(* Tests trace and span identifier generation.

   A generator fills its ring from the operating system guid service over ADS, so a fresh one
   has nothing to hand out until tick has been pumped for a few cycles. Every test that needs
   identifiers waits for that first refill before asserting anything about the bytes it gets
   back.

   Each test declares its generator in its own VAR_INST, next to the state machine that pumps
   it, so the ring a test reasons about is written down where the test reads it rather than in
   a list on the suite. Ring sizes are therefore chosen per test: most take a ring far larger
   than they draw from, so the seam never comes into it, while the wrap and capacity tests
   deliberately take the smallest ring the configuration allows, because a ring that small is
   the only one a test can drain often enough to lap. *)
FUNCTION_BLOCK FB_TestIdGenerator EXTENDS FB_TestSuite

THIS^.testRejectsInvalidConfiguration();
THIS^.testFailsBeforeTheFirstRefill();
THIS^.testGeneratesUniqueTraceIds();
THIS^.testGeneratesUniqueSpanIds();
THIS^.testDrawsAcrossTheWrap();
THIS^.testHonorsConfiguredCapacity();
THIS^.testGeneratesThroughTheBaseReference();
THIS^.testSeparateGeneratorsDoNotCollide();

(* TRUE when every byte in the buffer is zero, which is the identifier OTLP reads as absent. *)
METHOD _isZero : BOOL
VAR_INPUT
	pBytes: POINTER TO BYTE;
	nBytes: UDINT;
END_VAR
VAR
	_idx: UDINT;
END_VAR
_isZero := TRUE;

IF (pBytes = 0) OR_ELSE (nBytes = 0) THEN
	RETURN;
END_IF

FOR _idx := 0 TO nBytes - 1 DO
	IF pBytes[_idx] <> 0 THEN
		_isZero := FALSE;
		RETURN;
	END_IF
END_FOR
END_METHOD

(* Exercises the seam. A thirty two byte ring cannot hold eight identifiers at once, so the
   draws are spread over cycles and the read point laps the ring several times.

   Taking sixteen bytes and then eight moves the read point by twenty four, which lands it on
   every eight byte alignment in turn: some trace draws stop short of the end of the ring, one
   ends exactly on it, and one starts near the end and has to be stitched from both sides. A
   stitch that copied the wrong end, or re-read bytes already handed out, shows up here as a
   repeat among the samples. *)
METHOD testDrawsAcrossTheWrap : REFERENCE TO FB_Test

VAR CONSTANT
	MAX_CYCLES: UDINT := 60000;
	SAMPLES: UDINT := 8;
END_VAR

VAR_INST
	_generator: FB_IdGenerator(nTraceIds := 1, nSpanIds := 1);  // 24 bytes, which FB_Init rounds up to 32
	_cycles: UDINT;
	_state: USINT;
	_traceIdx: UDINT;
	_spanIdx: UDINT;
	_traceSamples: ARRAY [0..7, 0..15] OF BYTE;  // held across cycles, unlike the other suites
	_spanSamples: ARRAY [0..7, 0..7] OF BYTE;
END_VAR

VAR
	traceId: FB_TraceId;
	spanId: FB_SpanId;
	failureReason: E_IdGenFailureReason;
	tickSucceeded: BOOL;
	_i: UDINT;
	_j: UDINT;
END_VAR
TcUnit.TEST('testDrawsAcrossTheWrap');
	CASE _state OF
		0: // take whatever the ring can serve this cycle, however many laps that takes
			tickSucceeded := _generator.tick(failureReason=>failureReason);
			_cycles := _cycles + 1;
			IF NOT tickSucceeded THEN
				THIS^.AssertTrue(FALSE, 'Expected the guid service to refill the ring without error');
				_state := 255;
				TcUnit.TEST_FINISHED();
				RETURN;
			END_IF

			IF (_traceIdx < SAMPLES) AND_THEN _generator.generateTraceId(traceId:=traceId, failureReason=>failureReason) THEN
				MEMCPY(ADR(_traceSamples[_traceIdx, 0]), ADR(traceId.bytes), SIZEOF(traceId.bytes));
				_traceIdx := _traceIdx + 1;
			END_IF

			IF (_spanIdx < SAMPLES) AND_THEN _generator.generateSpanId(spanId:=spanId, failureReason=>failureReason) THEN
				MEMCPY(ADR(_spanSamples[_spanIdx, 0]), ADR(spanId.bytes), SIZEOF(spanId.bytes));
				_spanIdx := _spanIdx + 1;
			END_IF

			IF (_traceIdx >= SAMPLES) AND (_spanIdx >= SAMPLES) THEN
				_state := 10;
			ELSIF _cycles > MAX_CYCLES THEN
				THIS^.AssertTrue(FALSE, 'Expected a ring small enough to wrap to hand out its identifiers within MAX_CYCLES');
				_state := 255;
				TcUnit.TEST_FINISHED();
			END_IF
			RETURN;

		10:
			FOR _i := 0 TO 7 DO
				THIS^.AssertFalse(
					THIS^._isZero(pBytes:=ADR(_traceSamples[_i, 0]), nBytes:=TO_UDINT(SIZEOF(traceId.bytes))),
					'Expected no trace id drawn from a wrapping ring to be all zeroes'
				);
				THIS^.AssertFalse(
					THIS^._isZero(pBytes:=ADR(_spanSamples[_i, 0]), nBytes:=TO_UDINT(SIZEOF(spanId.bytes))),
					'Expected no span id drawn from a wrapping ring to be all zeroes'
				);

				FOR _j := 0 TO 7 DO
					IF _i <> _j THEN
						THIS^.AssertTrue(
							MEMCMP(ADR(_traceSamples[_i, 0]), ADR(_traceSamples[_j, 0]), SIZEOF(traceId.bytes)) <> 0,
							'Expected every trace id to differ, including the one stitched across the wrap'
						);
						THIS^.AssertTrue(
							MEMCMP(ADR(_spanSamples[_i, 0]), ADR(_spanSamples[_j, 0]), SIZEOF(spanId.bytes)) <> 0,
							'Expected every span id to differ, including the ones taken either side of the wrap'
						);
					END_IF
				END_FOR
			END_FOR

			_state := 255;
			TcUnit.TEST_FINISHED();
			RETURN;
	END_CASE
END_METHOD

(* A generator that has never been ticked holds no bytes. It has to say so, because the only
   thing it could hand out instead is the all zero identifier OTLP reads as absent. *)
METHOD testFailsBeforeTheFirstRefill : REFERENCE TO FB_Test

VAR_INST
	_generator: FB_IdGenerator(nTraceIds := 16, nSpanIds := 16);  // deliberately never ticked, so it stays empty
	_state: USINT;
END_VAR

VAR
	traceId: FB_TraceId;
	spanId: FB_SpanId;
	failureReason: E_IdGenFailureReason;
	success: BOOL;
END_VAR
TcUnit.TEST('testFailsBeforeTheFirstRefill');
	CASE _state OF
		0:
			THIS^.AssertTrue(_generator.configValid, 'Expected a generator with a ring to report a valid configuration');

			success := _generator.generateTraceId(traceId:=traceId, failureReason=>failureReason);
			THIS^.AssertFalse(success, 'Expected trace id generation to fail before the first refill');
			THIS^.AssertEquals_UDINT(
				TO_UDINT(E_IdGenFailureReason.NO_IDENTIFIERS_AVAILABLE),
				TO_UDINT(failureReason),
				'Expected an empty ring to report NO_IDENTIFIERS_AVAILABLE'
			);
			THIS^.AssertTrue(
				THIS^._isZero(pBytes:=ADR(traceId.bytes), nBytes:=TO_UDINT(SIZEOF(traceId.bytes))),
				'Expected a failed draw to leave the trace id untouched'
			);

			success := _generator.generateSpanId(spanId:=spanId, failureReason=>failureReason);
			THIS^.AssertFalse(success, 'Expected span id generation to fail before the first refill');
			THIS^.AssertEquals_UDINT(
				TO_UDINT(E_IdGenFailureReason.NO_IDENTIFIERS_AVAILABLE),
				TO_UDINT(failureReason),
				'Expected an empty ring to report NO_IDENTIFIERS_AVAILABLE'
			);
			THIS^.AssertTrue(
				THIS^._isZero(pBytes:=ADR(spanId.bytes), nBytes:=TO_UDINT(SIZEOF(spanId.bytes))),
				'Expected a failed draw to leave the span id untouched'
			);

			_state := 255;
			TcUnit.TEST_FINISHED();
	END_CASE
END_METHOD

(* Callers hold the generator as REFERENCE TO FB_IdGenerator_Base, so the abstract methods have
   to dispatch to the concrete ring. *)
METHOD testGeneratesThroughTheBaseReference : REFERENCE TO FB_Test

VAR CONSTANT
	MAX_CYCLES: UDINT := 60000;
END_VAR

VAR_INST
	_generator: FB_IdGenerator(nTraceIds := 16, nSpanIds := 16);
	_cycles: UDINT;
	_state: USINT;
END_VAR

VAR
	base: REFERENCE TO FB_IdGenerator_Base;
	traceId: FB_TraceId;
	spanId: FB_SpanId;
	failureReason: E_IdGenFailureReason;
	tickSucceeded: BOOL;
	success: BOOL;
END_VAR
TcUnit.TEST('testGeneratesThroughTheBaseReference');
	base REF= _generator;
	CASE _state OF
		0:
			THIS^.AssertTrue(__ISVALIDREF(base), 'Expected the base reference to be valid');
			_state := 10;
			RETURN;

		10: // pump through the base reference until the first refill lands
			tickSucceeded := base.tick(failureReason=>failureReason);
			_cycles := _cycles + 1;
			IF NOT tickSucceeded THEN
				THIS^.AssertTrue(FALSE, 'Expected tick to dispatch to the concrete generator without error');
				_state := 255;
				TcUnit.TEST_FINISHED();
				RETURN;
			END_IF

			success := base.generateTraceId(traceId:=traceId, failureReason=>failureReason);
			IF NOT success THEN
				IF _cycles > MAX_CYCLES THEN
					THIS^.AssertTrue(FALSE, 'Expected identifiers through the base reference within MAX_CYCLES');
					_state := 255;
					TcUnit.TEST_FINISHED();
				END_IF
				RETURN;
			END_IF

			THIS^.AssertFalse(
				THIS^._isZero(pBytes:=ADR(traceId.bytes), nBytes:=TO_UDINT(SIZEOF(traceId.bytes))),
				'Expected a non zero trace id through the base reference'
			);

			success := base.generateSpanId(spanId:=spanId, failureReason=>failureReason);
			THIS^.AssertTrue(success, 'Expected generateSpanId to dispatch to the concrete generator');
			THIS^.AssertFalse(
				THIS^._isZero(pBytes:=ADR(spanId.bytes), nBytes:=TO_UDINT(SIZEOF(spanId.bytes))),
				'Expected a non zero span id through the base reference'
			);

			_state := 255;
			TcUnit.TEST_FINISHED();
			RETURN;
	END_CASE
END_METHOD

(* The same requirement as for trace ids. A span id handed out twice makes two spans in the
   same trace indistinguishable. *)
METHOD testGeneratesUniqueSpanIds : REFERENCE TO FB_Test

VAR CONSTANT
	MAX_CYCLES: UDINT := 60000;
END_VAR

VAR_INST
	_generator: FB_IdGenerator(nTraceIds := 16, nSpanIds := 16);  // 384 bytes, so eight samples come out of one fill
	_cycles: UDINT;
	_state: USINT;
END_VAR

VAR
	spanId: FB_SpanId;
	samples: ARRAY [0..7, 0..7] OF BYTE;
	failureReason: E_IdGenFailureReason;
	tickSucceeded: BOOL;
	success: BOOL;
	_i: UDINT;
	_j: UDINT;
END_VAR
TcUnit.TEST('testGeneratesUniqueSpanIds');
	CASE _state OF
		0: // wait for the first refill before drawing the samples
			tickSucceeded := _generator.tick(failureReason=>failureReason);
			_cycles := _cycles + 1;
			IF NOT tickSucceeded THEN
				THIS^.AssertTrue(FALSE, 'Expected the guid service to refill the ring without error');
				_state := 255;
				TcUnit.TEST_FINISHED();
				RETURN;
			END_IF

			IF _generator.generateSpanId(spanId:=spanId, failureReason=>failureReason) THEN
				_state := 10;
			ELSIF _cycles > MAX_CYCLES THEN
				THIS^.AssertTrue(FALSE, 'Expected the first ring of span ids within MAX_CYCLES');
				_state := 255;
				TcUnit.TEST_FINISHED();
			END_IF
			RETURN;

		10: // a full ring holds forty eight span ids, so all eight samples come out of one fill
			FOR _i := 0 TO 7 DO
				success := _generator.generateSpanId(spanId:=spanId, failureReason=>failureReason);
				THIS^.AssertTrue(success, 'Expected every span id draw from a filled ring to succeed');
				THIS^.AssertEquals_UDINT(
					TO_UDINT(E_IdGenFailureReason.NA),
					TO_UDINT(failureReason),
					'Expected no failure reason alongside a successful draw'
				);
				THIS^.AssertFalse(
					THIS^._isZero(pBytes:=ADR(spanId.bytes), nBytes:=TO_UDINT(SIZEOF(spanId.bytes))),
					'Expected no span id to be all zeroes'
				);
				MEMCPY(ADR(samples[_i, 0]), ADR(spanId.bytes), SIZEOF(spanId.bytes));
			END_FOR

			FOR _i := 0 TO 7 DO
				FOR _j := 0 TO 7 DO
					IF _i <> _j THEN
						THIS^.AssertTrue(
							MEMCMP(ADR(samples[_i, 0]), ADR(samples[_j, 0]), SIZEOF(spanId.bytes)) <> 0,
							'Expected every span id to differ from every other'
						);
					END_IF
				END_FOR
			END_FOR

			_state := 255;
			TcUnit.TEST_FINISHED();
			RETURN;
	END_CASE
END_METHOD

(* Every draw has to be its own bytes. A trace id handed out twice merges two unrelated traces
   at the collector, which is worse than no trace at all. *)
METHOD testGeneratesUniqueTraceIds : REFERENCE TO FB_Test

VAR CONSTANT
	MAX_CYCLES: UDINT := 60000;
END_VAR

VAR_INST
	_generator: FB_IdGenerator(nTraceIds := 16, nSpanIds := 16);  // 384 bytes, so eight samples come out of one fill
	_cycles: UDINT;
	_state: USINT;
END_VAR

VAR
	traceId: FB_TraceId;
	samples: ARRAY [0..7, 0..15] OF BYTE;
	failureReason: E_IdGenFailureReason;
	tickSucceeded: BOOL;
	success: BOOL;
	_i: UDINT;
	_j: UDINT;
END_VAR
TcUnit.TEST('testGeneratesUniqueTraceIds');
	CASE _state OF
		0: // wait for the first refill before drawing the samples
			tickSucceeded := _generator.tick(failureReason=>failureReason);
			_cycles := _cycles + 1;
			IF NOT tickSucceeded THEN
				THIS^.AssertTrue(FALSE, 'Expected the guid service to refill the ring without error');
				_state := 255;
				TcUnit.TEST_FINISHED();
				RETURN;
			END_IF

			IF _generator.generateTraceId(traceId:=traceId, failureReason=>failureReason) THEN
				_state := 10;
			ELSIF _cycles > MAX_CYCLES THEN
				THIS^.AssertTrue(FALSE, 'Expected the first ring of trace ids within MAX_CYCLES');
				_state := 255;
				TcUnit.TEST_FINISHED();
			END_IF
			RETURN;

		10: // a full ring holds twenty four trace ids, so all eight samples come out of one fill
			FOR _i := 0 TO 7 DO
				success := _generator.generateTraceId(traceId:=traceId, failureReason=>failureReason);
				THIS^.AssertTrue(success, 'Expected every trace id draw from a filled ring to succeed');
				THIS^.AssertEquals_UDINT(
					TO_UDINT(E_IdGenFailureReason.NA),
					TO_UDINT(failureReason),
					'Expected no failure reason alongside a successful draw'
				);
				THIS^.AssertFalse(
					THIS^._isZero(pBytes:=ADR(traceId.bytes), nBytes:=TO_UDINT(SIZEOF(traceId.bytes))),
					'Expected no trace id to be all zeroes'
				);
				MEMCPY(ADR(samples[_i, 0]), ADR(traceId.bytes), SIZEOF(traceId.bytes));
			END_FOR

			FOR _i := 0 TO 7 DO
				FOR _j := 0 TO 7 DO
					IF _i <> _j THEN
						THIS^.AssertTrue(
							MEMCMP(ADR(samples[_i, 0]), ADR(samples[_j, 0]), SIZEOF(traceId.bytes)) <> 0,
							'Expected every trace id to differ from every other'
						);
					END_IF
				END_FOR
			END_FOR

			_state := 255;
			TcUnit.TEST_FINISHED();
			RETURN;
	END_CASE
END_METHOD

(* One trace id and one span id is twenty four bytes, which FB_Init rounds up to thirty two
   because the guid service will not write anything narrower than a whole guid. A full ring is
   therefore exactly two trace ids wide, and no amount of refilling grows it past that. *)
METHOD testHonorsConfiguredCapacity : REFERENCE TO FB_Test

VAR CONSTANT
	MAX_CYCLES: UDINT := 60000;
	MAX_DRAWS: UDINT := 16;  // comfortably more than a thirty two byte ring could ever serve
	EXPECTED_TRACE_IDS: UDINT := 2;
END_VAR

VAR_INST
	_generator: FB_IdGenerator(nTraceIds := 1, nSpanIds := 1);  // the shortest ring the configuration allows
	_cycles: UDINT;
	_state: USINT;
	_best: UDINT;  // the most trace ids any single drain has yielded
END_VAR

VAR
	traceId: FB_TraceId;
	failureReason: E_IdGenFailureReason;
	tickSucceeded: BOOL;
	drawn: UDINT;
	_i: UDINT;
END_VAR
TcUnit.TEST('testHonorsConfiguredCapacity');
	CASE _state OF
		0: // drain the ring dry every cycle, so the best any one drain manages is one full ring
			tickSucceeded := _generator.tick(failureReason=>failureReason);
			_cycles := _cycles + 1;
			IF NOT tickSucceeded THEN
				THIS^.AssertTrue(FALSE, 'Expected the guid service to refill the ring without error');
				_state := 255;
				TcUnit.TEST_FINISHED();
				RETURN;
			END_IF

			drawn := 0;
			FOR _i := 1 TO MAX_DRAWS DO
				IF NOT _generator.generateTraceId(traceId:=traceId, failureReason=>failureReason) THEN
					EXIT;
				END_IF
				drawn := drawn + 1;
			END_FOR

			THIS^.AssertTrue(
				drawn <= EXPECTED_TRACE_IDS,
				'Expected a refill never to serve more than the configured ring holds'
			);
			THIS^.AssertEquals_UDINT(
				TO_UDINT(E_IdGenFailureReason.NO_IDENTIFIERS_AVAILABLE),
				TO_UDINT(failureReason),
				'Expected the draw that emptied the ring to report NO_IDENTIFIERS_AVAILABLE'
			);

			IF drawn > _best THEN
				_best := drawn;
			END_IF

			IF _best >= EXPECTED_TRACE_IDS THEN
				_state := 10;
			ELSIF _cycles > MAX_CYCLES THEN
				THIS^.AssertTrue(FALSE, 'Expected the ring to fill to its configured length within MAX_CYCLES');
				_state := 255;
				TcUnit.TEST_FINISHED();
			END_IF
			RETURN;

		10:
			THIS^.AssertEquals_UDINT(
				EXPECTED_TRACE_IDS,
				_best,
				'Expected a twenty four byte request to become a thirty two byte ring'
			);
			_state := 255;
			TcUnit.TEST_FINISHED();
			RETURN;
	END_CASE
END_METHOD

(* A generator asked for no identifiers never allocates a ring, so every entry point has to say
   so rather than read through a null pointer. *)
METHOD testRejectsInvalidConfiguration : REFERENCE TO FB_Test

VAR_INST
	_generator: FB_IdGenerator(nTraceIds := 0, nSpanIds := 0);  // asks for nothing, so no ring is allocated
	_state: USINT;
END_VAR

VAR
	traceId: FB_TraceId;
	spanId: FB_SpanId;
	failureReason: E_IdGenFailureReason;
	success: BOOL;
END_VAR
TcUnit.TEST('testRejectsInvalidConfiguration');
	CASE _state OF
		0:
			THIS^.AssertFalse(_generator.configValid, 'Expected a generator with no ring to report an invalid configuration');

			success := _generator.tick(failureReason=>failureReason);
			THIS^.AssertFalse(success, 'Expected tick to fail when no ring was allocated');
			THIS^.AssertEquals_UDINT(
				TO_UDINT(E_IdGenFailureReason.INVALID_CONFIGUATION),
				TO_UDINT(failureReason),
				'Expected tick to report INVALID_CONFIGUATION'
			);

			success := _generator.generateTraceId(traceId:=traceId, failureReason=>failureReason);
			THIS^.AssertFalse(success, 'Expected trace id generation to fail when no ring was allocated');
			THIS^.AssertEquals_UDINT(
				TO_UDINT(E_IdGenFailureReason.INVALID_CONFIGUATION),
				TO_UDINT(failureReason),
				'Expected a missing ring to be reported as a configuration mistake, not an empty ring'
			);

			success := _generator.generateSpanId(spanId:=spanId, failureReason=>failureReason);
			THIS^.AssertFalse(success, 'Expected span id generation to fail when no ring was allocated');
			THIS^.AssertEquals_UDINT(
				TO_UDINT(E_IdGenFailureReason.INVALID_CONFIGUATION),
				TO_UDINT(failureReason),
				'Expected a missing ring to be reported as a configuration mistake, not an empty ring'
			);

			_state := 255;
			TcUnit.TEST_FINISHED();
	END_CASE
END_METHOD

(* Two generators built in the same cycle must not emit the same identifiers, or two providers
   on one PLC would report traces the collector cannot tell apart. *)
METHOD testSeparateGeneratorsDoNotCollide : REFERENCE TO FB_Test

VAR CONSTANT
	MAX_CYCLES: UDINT := 60000;
END_VAR

VAR_INST
	_generatorA: FB_IdGenerator(nTraceIds := 16, nSpanIds := 16);
	_generatorB: FB_IdGenerator(nTraceIds := 16, nSpanIds := 16);
	_cycles: UDINT;
	_state: USINT;
END_VAR

VAR
	traceIdA: FB_TraceId;
	traceIdB: FB_TraceId;
	spanIdA: FB_SpanId;
	spanIdB: FB_SpanId;
	failureReason: E_IdGenFailureReason;
	tickSucceededA: BOOL;
	tickSucceededB: BOOL;
	drewA: BOOL;
	drewB: BOOL;
	success: BOOL;
END_VAR
TcUnit.TEST('testSeparateGeneratorsDoNotCollide');
	CASE _state OF
		0: // pump both rings until they can each serve in the same cycle
			tickSucceededA := _generatorA.tick(failureReason=>failureReason);
			tickSucceededB := _generatorB.tick(failureReason=>failureReason);
			_cycles := _cycles + 1;
			IF NOT (tickSucceededA AND tickSucceededB) THEN
				THIS^.AssertTrue(FALSE, 'Expected both generators to refill without error');
				_state := 255;
				TcUnit.TEST_FINISHED();
				RETURN;
			END_IF

			// both are drawn unconditionally, so neither ring is drained ahead of the other
			drewA := _generatorA.generateTraceId(traceId:=traceIdA, failureReason=>failureReason);
			drewB := _generatorB.generateTraceId(traceId:=traceIdB, failureReason=>failureReason);
			IF NOT (drewA AND drewB) THEN
				IF _cycles > MAX_CYCLES THEN
					THIS^.AssertTrue(FALSE, 'Expected both generators to fill within MAX_CYCLES');
					_state := 255;
					TcUnit.TEST_FINISHED();
				END_IF
				RETURN;
			END_IF

			THIS^.AssertTrue(
				MEMCMP(ADR(traceIdA.bytes), ADR(traceIdB.bytes), SIZEOF(traceIdA.bytes)) <> 0,
				'Expected two generators to produce different trace ids'
			);

			success := _generatorA.generateSpanId(spanId:=spanIdA, failureReason=>failureReason);
			THIS^.AssertTrue(success, 'Expected the first generator to serve a span id from a filled ring');
			success := _generatorB.generateSpanId(spanId:=spanIdB, failureReason=>failureReason);
			THIS^.AssertTrue(success, 'Expected the second generator to serve a span id from a filled ring');
			THIS^.AssertTrue(
				MEMCMP(ADR(spanIdA.bytes), ADR(spanIdB.bytes), SIZEOF(spanIdA.bytes)) <> 0,
				'Expected two generators to produce different span ids'
			);

			_state := 255;
			TcUnit.TEST_FINISHED();
			RETURN;
	END_CASE
END_METHOD

END_FUNCTION_BLOCK

(* stored: Version 1.1.0.1
   POU FB_TestIdGenerator: Id {8b541683-370a-4944-9efb-d4dbe8f57299}, SpecialFunc None
   Method _isZero: Id {5705a4f9-bf6a-4d55-849b-bcecacb7cf3f}
   Method testDrawsAcrossTheWrap: Id {9792fca8-fa0f-415e-a698-2a0efab33a17}
   Method testFailsBeforeTheFirstRefill: Id {fa5f5605-0d88-4c65-a08f-8e7758eb0e3c}
   Method testGeneratesThroughTheBaseReference: Id {368b4998-ac3d-460a-b25b-6f8821b1bb3e}
   Method testGeneratesUniqueSpanIds: Id {e90fe6c4-350b-4279-9671-f4dbf9765e7e}
   Method testGeneratesUniqueTraceIds: Id {9de941f7-0da5-48b8-8337-8561a784824b}
   Method testHonorsConfiguredCapacity: Id {436d3595-2483-4d76-bfbf-a554ad7ac412}
   Method testRejectsInvalidConfiguration: Id {7bd81400-5827-4199-b8a2-f5efaa1ca167}
   Method testSeparateGeneratorsDoNotCollide: Id {d1410e95-1088-446d-9d92-44e00dfb0300} *)
